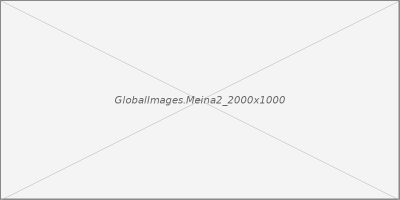
VISUALIZATION V_NCIMeina2_2000x1000  // 400x200
VAR_IN_OUT
	HMI : ST_PackMLBaseModule_HMI;
	HMI_GantryXYZ : ST_GantryXYZ_HMI;
	HMI_Recipe : ST_RecipeBuilder_HMI;
END_VAR
    RoundedRectangle (0,0 400x200)
    Image (0,0 400x200), image: GlobalImages.Meina2_2000x1000
END_VISUALIZATION

(* stored: Version 1.1.0.1, ProductVersion 3.1.4024.15
   Visu V_NCIMeina2_2000x1000: Id {f140fc45-fca9-4039-8c48-b52e58f74615} *)
